(* IEC 61131-3 sources: plc-st-test/packages/cli/test/fixtures/ambiguous/Tests, 1 file *)

(* ---- TEST_Any.st ---- *)
FUNCTION_BLOCK TEST_Any
METHOD Test_Nothing
  ASSERT_TRUE(TRUE);
END_METHOD
END_FUNCTION_BLOCK
